FUNCTION FC 1 : VOID
BEGIN
NETWORK
      CU C 300
END_FUNCTION
